(* IEC 61131-3 sources: stc/stdlib/vendor/beckhoff, 10 files *)

(* ---- common_types.st ---- *)
(* Common types used across Beckhoff TwinCAT 3 libraries *)
(* Stub declarations for stc type-checking. No implementation bodies. *)

(* AXIS_REF -- Opaque axis reference structure used by all MC_* blocks *)
TYPE AXIS_REF :
STRUCT
    NcToPlc     : DINT;
    PlcToNc     : DINT;
END_STRUCT
END_TYPE

(* MC_Direction -- Motion direction for MC_MoveAbsolute, MC_MoveVelocity *)
TYPE MC_Direction : (
    mcPositiveDirection,
    mcNegativeDirection,
    mcCurrentDirection,
    mcShortestWay
);
END_TYPE

(* T_AmsNetId -- AMS Net ID string for ADS communication *)
TYPE T_AmsNetId : STRING(23); END_TYPE

(* T_AmsPort -- AMS port number *)
TYPE T_AmsPort : UINT; END_TYPE

(* T_MaxString -- General-purpose maximum-length string *)
TYPE T_MaxString : STRING(255); END_TYPE

(* E_OpenPath -- File open path options for FB_FileOpen *)
TYPE E_OpenPath : (
    PATH_GENERIC,
    PATH_BOOTPATH,
    PATH_BOOTPRJPATH
);
END_TYPE

(* PVOID -- untyped address. TwinCAT defines PVOID as UXINT (ULINT on 64-bit,
   UDINT on 32-bit). stc declares it as POINTER TO BYTE (locked Phase 21
   decision). Phase 22 must make ADR(...) results and any POINTER TO <T>
   assignable to PVOID. *)
TYPE PVOID : POINTER TO BYTE; END_TYPE

(* Platform-width integer aliases (TwinCAT PLC manual 16.5.11), 64-bit sizes *)
TYPE __XWORD : LWORD; END_TYPE

TYPE XWORD : LWORD; END_TYPE

TYPE UXINT : ULINT; END_TYPE

TYPE __UXINT : ULINT; END_TYPE

TYPE XINT : LINT; END_TYPE

TYPE __XINT : LINT; END_TYPE

(* AMSPORT -- AMS port number (Tc2_System alias) *)
TYPE AMSPORT : UINT; END_TYPE

(* ---- tc3_ipcdiag.st ---- *)
(* Tc3_IPCDiag -- placeholder stub *)
(* No symbols from this library are used by sildarvinnsla; the file is
   present so the library reference resolves. The marker type below keeps
   the one-declaration-per-stub rule and is not a Beckhoff symbol. *)

TYPE T_Tc3IPCDiagStubMarker : BOOL; END_TYPE

(* ---- tc3_module.st ---- *)
(* Tc3_Module -- placeholder stub *)
(* No symbols from this library are used by sildarvinnsla; the file is
   present so the library reference resolves. The marker type below keeps
   the one-declaration-per-stub rule and is not a Beckhoff symbol. *)

TYPE T_Tc3ModuleStubMarker : BOOL; END_TYPE

(* ---- tc2_ethercat.st ---- *)
(* Tc2_EtherCAT -- EtherCAT diagnostics and mailbox function blocks *)
(* Stub declarations for stc type-checking. No implementation bodies. *)
(* Source: TwinCAT 3 PLC Lib Tc2_EtherCAT manual v1.10.0. *)
(* E_EcSlaveState, EcDiagParam and FB_EcDeviceDiag are deliberately NOT
   declared here: they are SVNCoreComponents declarations, not Beckhoff
   ones, and must resolve from that library. *)

TYPE E_EcAdressingType : (
    eAdressingType_AutoInc := 1,
    eAdressingType_Fixed,
    eAdressingType_Broadcast
);
END_TYPE

TYPE ST_EcSlaveState :
STRUCT
    deviceState     : BYTE;
    linkState       : BYTE;
END_STRUCT
END_TYPE

TYPE ST_EcCrcError :
STRUCT
    portA           : UDINT;
    portB           : UDINT;
    portC           : UDINT;
END_STRUCT
END_TYPE

TYPE ST_EcCrcErrorEx :
STRUCT
    portA           : UDINT;
    portB           : UDINT;
    portC           : UDINT;
    portD           : UDINT;
END_STRUCT
END_TYPE

(* Global constants, section 14.1 (subset) *)
VAR_GLOBAL CONSTANT
    EC_AMSPORT_MASTER               : UINT := 16#FFFF;
    EC_MAX_SLAVES                   : UINT := 16#FFFF;
    EC_DEVICE_STATE_MASK            : BYTE := 16#0F;
    EC_DEVICE_STATE_INIT            : BYTE := 16#01;
    EC_DEVICE_STATE_PREOP           : BYTE := 16#02;
    EC_DEVICE_STATE_BOOTSTRAP       : BYTE := 16#03;
    EC_DEVICE_STATE_SAFEOP          : BYTE := 16#04;
    EC_DEVICE_STATE_OP              : BYTE := 16#08;
    EC_DEVICE_STATE_ERROR           : BYTE := 16#10;
    EC_DEVICE_STATE_INVALID_VPRS    : BYTE := 16#20;
    EC_DEVICE_STATE_INITCMD_ERROR   : BYTE := 16#40;
    EC_LINK_STATE_OK                : BYTE := 16#00;
    EC_LINK_STATE_NOT_PRESENT       : BYTE := 16#01;
    EC_LINK_STATE_LINK_WITHOUT_COMM : BYTE := 16#02;
    EC_LINK_STATE_MISSING_LINK      : BYTE := 16#04;
    EC_LINK_STATE_ADDITIONAL_LINK   : BYTE := 16#08;
    EC_LINK_STATE_PORT_A            : BYTE := 16#10;
    EC_LINK_STATE_PORT_B            : BYTE := 16#20;
    EC_LINK_STATE_PORT_C            : BYTE := 16#40;
    EC_LINK_STATE_PORT_D            : BYTE := 16#80;
END_VAR

(* Section 3.2 *)
FUNCTION_BLOCK FB_EcPhysicalWriteCmd
VAR_INPUT
    sNetId          : T_AmsNetId;
    adp             : UINT;
    ado             : UINT;
    len             : UDINT;
    eType           : E_EcAdressingType := eAdressingType_Fixed;
    pSrcBuf         : PVOID;
    bExecute        : BOOL;
    tTimeout        : TIME := DEFAULT_ADS_TIMEOUT;
END_VAR
VAR_OUTPUT
    bBusy           : BOOL;
    bError          : BOOL;
    nErrId          : UDINT;
    wkc             : UINT;
END_VAR
END_FUNCTION_BLOCK

(* Section 4.3 *)
FUNCTION_BLOCK FB_EcGetAllSlaveAddr
VAR_INPUT
    sNetId          : T_AmsNetId;
    pAddrBuf        : POINTER TO ARRAY[0..EC_MAX_SLAVES] OF UINT;
    cbBufLen        : UDINT;
    bExecute        : BOOL;
    tTimeout        : TIME := DEFAULT_ADS_TIMEOUT;
END_VAR
VAR_OUTPUT
    bBusy           : BOOL;
    bError          : BOOL;
    nErrId          : UDINT;
    nSlaves         : UINT;
END_VAR
END_FUNCTION_BLOCK

(* Section 4.4 *)
FUNCTION_BLOCK FB_EcGetAllSlaveCrcErrors
VAR_INPUT
    sNetId          : T_AmsNetId;
    pCrcErrorBuf    : POINTER TO ARRAY[0..EC_MAX_SLAVES] OF DWORD;
    cbBufLen        : UDINT;
    bExecute        : BOOL;
    tTimeout        : TIME := DEFAULT_ADS_TIMEOUT;
END_VAR
VAR_OUTPUT
    bBusy           : BOOL;
    bError          : BOOL;
    nErrId          : UDINT;
    nSlaves         : UINT;
END_VAR
END_FUNCTION_BLOCK

(* Section 4.12 *)
FUNCTION_BLOCK FB_EcGetSlaveCrcError
VAR_INPUT
    sNetId          : T_AmsNetId;
    nSlaveAddr      : UINT;
    bExecute        : BOOL;
    tTimeout        : TIME := DEFAULT_ADS_TIMEOUT;
END_VAR
VAR_OUTPUT
    bBusy           : BOOL;
    bError          : BOOL;
    nErrId          : UDINT;
    crcError        : ST_EcCrcError;
END_VAR
END_FUNCTION_BLOCK

(* Section 4.13 (tTimeout has no default in the manual) *)
FUNCTION_BLOCK FB_EcGetSlaveCrcErrorEx
VAR_INPUT
    sNetId          : T_AmsNetId;
    nSlaveAddr      : UINT;
    bExecute        : BOOL;
    tTimeout        : TIME;
END_VAR
VAR_OUTPUT
    bBusy           : BOOL;
    bError          : BOOL;
    nErrId          : UDINT;
    CrcError        : ST_EcCrcErrorEx;
END_VAR
END_FUNCTION_BLOCK

(* Section 5.1 *)
FUNCTION_BLOCK FB_EcGetAllSlaveStates
VAR_INPUT
    sNetId          : T_AmsNetId;
    pStateBuf       : POINTER TO ARRAY[0..EC_MAX_SLAVES] OF ST_EcSlaveState;
    cbBufLen        : UDINT;
    bExecute        : BOOL;
    tTimeout        : TIME := DEFAULT_ADS_TIMEOUT;
END_VAR
VAR_OUTPUT
    bBusy           : BOOL;
    bError          : BOOL;
    nErrId          : UDINT;
    nSlaves         : UINT;
END_VAR
END_FUNCTION_BLOCK

(* Section 5.3 *)
FUNCTION_BLOCK FB_EcGetMasterState
VAR_INPUT
    sNetId          : T_AmsNetId;
    bExecute        : BOOL;
    tTimeout        : TIME := DEFAULT_ADS_TIMEOUT;
END_VAR
VAR_OUTPUT
    bBusy           : BOOL;
    bError          : BOOL;
    nErrId          : UDINT;
    state           : WORD;
END_VAR
END_FUNCTION_BLOCK

(* Section 5.4 *)
FUNCTION_BLOCK FB_EcGetSlaveState
VAR_INPUT
    sNetId          : T_AmsNetId;
    nSlaveAddr      : UINT;
    bExecute        : BOOL;
    tTimeout        : TIME := DEFAULT_ADS_TIMEOUT;
END_VAR
VAR_OUTPUT
    bBusy           : BOOL;
    bError          : BOOL;
    nErrId          : UDINT;
    state           : ST_EcSlaveState;
END_VAR
END_FUNCTION_BLOCK

(* Section 5.9 *)
FUNCTION_BLOCK FB_EcSetSlaveState
VAR_INPUT
    sNetId          : T_AmsNetId;
    nSlaveAddr      : UINT;
    bExecute        : BOOL;
    tTimeout        : TIME := T#10S;
    reqState        : WORD;
END_VAR
VAR_OUTPUT
    bBusy           : BOOL;
    bError          : BOOL;
    nErrId          : UDINT;
    currState       : ST_EcSlaveState;
END_VAR
END_FUNCTION_BLOCK

(* Section 7.1 (Beckhoff also spells it FB_EcCoeSdoRead; names are case-insensitive) *)
FUNCTION_BLOCK FB_EcCoESdoRead
VAR_INPUT
    sNetId          : T_AmsNetId;
    nSlaveAddr      : UINT;
    nSubIndex       : BYTE;
    nIndex          : WORD;
    pDstBuf         : PVOID;
    cbBufLen        : UDINT;
    bExecute        : BOOL;
    tTimeout        : TIME := DEFAULT_ADS_TIMEOUT;
END_VAR
VAR_OUTPUT
    bBusy           : BOOL;
    bError          : BOOL;
    nErrId          : UDINT;
    cbRead          : UDINT;
END_VAR
END_FUNCTION_BLOCK

(* Section 7.3 *)
FUNCTION_BLOCK FB_EcCoESdoWrite
VAR_INPUT
    sNetId          : T_AmsNetId;
    nSlaveAddr      : UINT;
    nSubIndex       : BYTE;
    nIndex          : WORD;
    pSrcBuf         : PVOID;
    cbBufLen        : UDINT;
    bExecute        : BOOL;
    tTimeout        : TIME := DEFAULT_ADS_TIMEOUT;
END_VAR
VAR_OUTPUT
    bBusy           : BOOL;
    bError          : BOOL;
    nErrId          : UDINT;
END_VAR
END_FUNCTION_BLOCK

(* ---- tc2_mc2.st ---- *)
(* Tc2_MC2 -- PLCopen Motion Control function blocks for Beckhoff TwinCAT 3 *)
(* Stub declarations for stc type-checking. No implementation bodies. *)

FUNCTION_BLOCK MC_Power
VAR_INPUT
    Axis            : AXIS_REF;
    Enable          : BOOL;
    Enable_Positive : BOOL;
    Enable_Negative : BOOL;
    Override_V      : LREAL := 100.0;
END_VAR
VAR_OUTPUT
    Status      : BOOL;
    Busy        : BOOL;
    Active      : BOOL;
    Error       : BOOL;
    ErrorID     : UDINT;
END_VAR
END_FUNCTION_BLOCK

FUNCTION_BLOCK MC_MoveAbsolute
VAR_INPUT
    Axis            : AXIS_REF;
    Execute         : BOOL;
    Position        : LREAL;
    Velocity        : LREAL;
    Acceleration    : LREAL;
    Deceleration    : LREAL;
    Jerk            : LREAL;
    Direction       : MC_Direction;
END_VAR
VAR_OUTPUT
    Done            : BOOL;
    Busy            : BOOL;
    Active          : BOOL;
    CommandAborted  : BOOL;
    Error           : BOOL;
    ErrorID         : UDINT;
END_VAR
END_FUNCTION_BLOCK

FUNCTION_BLOCK MC_MoveRelative
VAR_INPUT
    Axis            : AXIS_REF;
    Execute         : BOOL;
    Distance        : LREAL;
    Velocity        : LREAL;
    Acceleration    : LREAL;
    Deceleration    : LREAL;
    Jerk            : LREAL;
END_VAR
VAR_OUTPUT
    Done            : BOOL;
    Busy            : BOOL;
    Active          : BOOL;
    CommandAborted  : BOOL;
    Error           : BOOL;
    ErrorID         : UDINT;
END_VAR
END_FUNCTION_BLOCK

FUNCTION_BLOCK MC_MoveVelocity
VAR_INPUT
    Axis            : AXIS_REF;
    Execute         : BOOL;
    Velocity        : LREAL;
    Acceleration    : LREAL;
    Deceleration    : LREAL;
    Jerk            : LREAL;
    Direction       : MC_Direction;
END_VAR
VAR_OUTPUT
    InVelocity      : BOOL;
    Busy            : BOOL;
    Active          : BOOL;
    CommandAborted  : BOOL;
    Error           : BOOL;
    ErrorID         : UDINT;
END_VAR
END_FUNCTION_BLOCK

FUNCTION_BLOCK MC_Stop
VAR_INPUT
    Axis            : AXIS_REF;
    Execute         : BOOL;
    Deceleration    : LREAL;
    Jerk            : LREAL;
END_VAR
VAR_OUTPUT
    Done            : BOOL;
    Busy            : BOOL;
    Active          : BOOL;
    CommandAborted  : BOOL;
    Error           : BOOL;
    ErrorID         : UDINT;
END_VAR
END_FUNCTION_BLOCK

FUNCTION_BLOCK MC_Home
VAR_INPUT
    Axis            : AXIS_REF;
    Execute         : BOOL;
    Position        : LREAL;
END_VAR
VAR_OUTPUT
    Done            : BOOL;
    Busy            : BOOL;
    Active          : BOOL;
    CommandAborted  : BOOL;
    Error           : BOOL;
    ErrorID         : UDINT;
END_VAR
END_FUNCTION_BLOCK

FUNCTION_BLOCK MC_Reset
VAR_INPUT
    Axis            : AXIS_REF;
    Execute         : BOOL;
END_VAR
VAR_OUTPUT
    Done            : BOOL;
    Busy            : BOOL;
    Error           : BOOL;
    ErrorID         : UDINT;
END_VAR
END_FUNCTION_BLOCK

FUNCTION_BLOCK MC_ReadActualPosition
VAR_INPUT
    Axis            : AXIS_REF;
    Enable          : BOOL;
END_VAR
VAR_OUTPUT
    Valid           : BOOL;
    Busy            : BOOL;
    Error           : BOOL;
    ErrorID         : UDINT;
    Position        : LREAL;
END_VAR
END_FUNCTION_BLOCK

FUNCTION_BLOCK MC_ReadActualVelocity
VAR_INPUT
    Axis            : AXIS_REF;
    Enable          : BOOL;
END_VAR
VAR_OUTPUT
    Valid           : BOOL;
    Busy            : BOOL;
    Error           : BOOL;
    ErrorID         : UDINT;
    ActualVelocity  : LREAL;
END_VAR
END_FUNCTION_BLOCK

FUNCTION_BLOCK MC_ReadStatus
VAR_INPUT
    Axis            : AXIS_REF;
    Enable          : BOOL;
END_VAR
VAR_OUTPUT
    Valid               : BOOL;
    Busy                : BOOL;
    Error               : BOOL;
    ErrorID             : UDINT;
    ErrorStop           : BOOL;
    Disabled            : BOOL;
    Stopping            : BOOL;
    StandStill          : BOOL;
    DiscreteMotion      : BOOL;
    ContinuousMotion    : BOOL;
    SynchronizedMotion  : BOOL;
    Homing              : BOOL;
END_VAR
END_FUNCTION_BLOCK

(* ---- tc2_modbussrv.st ---- *)
(* Tc2_ModbusSrv -- Modbus TCP client function blocks (TF6250) *)
(* Stub declarations for stc type-checking. No implementation bodies. *)
(* Source: TF6250 TC3 Modbus TCP manual section 6.1.2. Section 6.1 states the
   Modbus functions are implemented in the PLC library Tc2_ModbusSrv, which is
   the library name TwinCAT projects reference, so the client FBs live here. *)

VAR_GLOBAL CONSTANT
    MODBUS_TCP_PORT : UINT := 502;      (* value assumed: Modbus TCP standard port *)
END_VAR

(* Modbus function 1 *)
FUNCTION_BLOCK FB_MBReadCoils
VAR_INPUT
    sIPAddr         : STRING(15);
    nTCPPort        : UINT := MODBUS_TCP_PORT;
    nUnitID         : BYTE := 16#FF;
    nQuantity       : WORD;
    nMBAddr         : WORD;
    cbLength        : UDINT;
    pDestAddr       : POINTER TO BYTE;
    bExecute        : BOOL;
    tTimeout        : TIME;
END_VAR
VAR_OUTPUT
    bBUSY           : BOOL;
    bError          : BOOL;
    nErrId          : UDINT;
    cbRead          : UDINT;
END_VAR
END_FUNCTION_BLOCK

(* Modbus function 2 *)
FUNCTION_BLOCK FB_MBReadInputs
VAR_INPUT
    sIPAddr         : STRING(15);
    nTCPPort        : UINT := MODBUS_TCP_PORT;
    nUnitID         : BYTE := 16#FF;
    nQuantity       : WORD;
    nMBAddr         : WORD;
    cbLength        : UDINT;
    pDestAddr       : POINTER TO BYTE;
    bExecute        : BOOL;
    tTimeout        : TIME;
END_VAR
VAR_OUTPUT
    bBUSY           : BOOL;
    bError          : BOOL;
    nErrId          : UDINT;
    cbRead          : UDINT;
END_VAR
END_FUNCTION_BLOCK

(* Modbus function 3 *)
FUNCTION_BLOCK FB_MBReadRegs
VAR_INPUT
    sIPAddr         : STRING(15);
    nTCPPort        : UINT := MODBUS_TCP_PORT;
    nUnitID         : BYTE := 16#FF;
    nQuantity       : WORD;
    nMBAddr         : WORD;
    cbLength        : UDINT;
    pDestAddr       : POINTER TO BYTE;
    bExecute        : BOOL;
    tTimeout        : TIME;
END_VAR
VAR_OUTPUT
    bBUSY           : BOOL;
    bError          : BOOL;
    nErrId          : UDINT;
    cbRead          : UDINT;
END_VAR
END_FUNCTION_BLOCK

(* Modbus function 4 *)
FUNCTION_BLOCK FB_MBReadInputRegs
VAR_INPUT
    sIPAddr         : STRING(15);
    nTCPPort        : UINT := MODBUS_TCP_PORT;
    nUnitID         : BYTE := 16#FF;
    nQuantity       : WORD;
    nMBAddr         : WORD;
    cbLength        : UDINT;
    pDestAddr       : POINTER TO BYTE;
    bExecute        : BOOL;
    tTimeout        : TIME;
END_VAR
VAR_OUTPUT
    bBUSY           : BOOL;
    bError          : BOOL;
    nErrId          : UDINT;
    cbRead          : UDINT;
END_VAR
END_FUNCTION_BLOCK

(* Modbus function 5 *)
FUNCTION_BLOCK FB_MBWriteSingleCoil
VAR_INPUT
    sIPAddr         : STRING(15);
    nTCPPort        : UINT := MODBUS_TCP_PORT;
    nUnitID         : BYTE := 16#FF;
    nMBAddr         : WORD;
    nValue          : WORD;
    bExecute        : BOOL;
    tTimeout        : TIME;
END_VAR
VAR_OUTPUT
    bBUSY           : BOOL;
    bError          : BOOL;
    nErrId          : UDINT;
END_VAR
END_FUNCTION_BLOCK

(* Modbus function 6 *)
FUNCTION_BLOCK FB_MBWriteSingleReg
VAR_INPUT
    sIPAddr         : STRING(15);
    nTCPPort        : UINT := MODBUS_TCP_PORT;
    nUnitID         : BYTE := 16#FF;
    nMBAddr         : WORD;
    nValue          : WORD;
    bExecute        : BOOL;
    tTimeout        : TIME;
END_VAR
VAR_OUTPUT
    bBUSY           : BOOL;
    bError          : BOOL;
    nErrId          : UDINT;
END_VAR
END_FUNCTION_BLOCK

(* Modbus function 15 *)
FUNCTION_BLOCK FB_MBWriteCoils
VAR_INPUT
    sIPAddr         : STRING(15);
    nTCPPort        : UINT := MODBUS_TCP_PORT;
    nUnitID         : BYTE := 16#FF;
    nQuantity       : WORD;
    nMBAddr         : WORD;
    cbLength        : UDINT;
    pSrcAddr        : POINTER TO BYTE;
    bExecute        : BOOL;
    tTimeout        : TIME;
END_VAR
VAR_OUTPUT
    bBUSY           : BOOL;
    bError          : BOOL;
    nErrId          : UDINT;
END_VAR
END_FUNCTION_BLOCK

(* Modbus function 16 *)
FUNCTION_BLOCK FB_MBWriteRegs
VAR_INPUT
    sIPAddr         : STRING(15);
    nTCPPort        : UINT := MODBUS_TCP_PORT;
    nUnitID         : BYTE := 16#FF;
    nQuantity       : WORD;
    nMBAddr         : WORD;
    cbLength        : UDINT;
    pSrcAddr        : POINTER TO BYTE;
    bExecute        : BOOL;
    tTimeout        : TIME;
END_VAR
VAR_OUTPUT
    bBUSY           : BOOL;
    bError          : BOOL;
    nErrId          : UDINT;
END_VAR
END_FUNCTION_BLOCK

(* Modbus function 23 *)
FUNCTION_BLOCK FB_MBReadWriteRegs
VAR_INPUT
    sIPAddr         : STRING(15);
    nTCPPort        : UINT := MODBUS_TCP_PORT;
    nUnitID         : BYTE := 16#FF;
    nReadQuantity   : WORD;
    nMBReadAddr     : WORD;
    nWriteQuantity  : WORD;
    nMBWriteAddr    : WORD;
    cbDestLength    : UDINT;
    pDestAddr       : POINTER TO BYTE;
    cbSrcLength     : UDINT;
    pSrcAddr        : POINTER TO BYTE;
    bExecute        : BOOL;
    tTimeout        : TIME;
END_VAR
VAR_OUTPUT
    bBUSY           : BOOL;
    bError          : BOOL;
    nErrId          : UDINT;
    cbRead          : UDINT;
END_VAR
END_FUNCTION_BLOCK

(* ---- tc2_serialcom.st ---- *)
(* Tc2_SerialCom -- serial communication function blocks (TF6340) *)
(* Stub declarations for stc type-checking. No implementation bodies. *)
(* Source: TF6340 TC3 Serial Communication manual section 5. The real type
   names are ComBuffer, ComSerialLineMode_t and ComError_t (ST_ComBuffer and
   E_ComMode do not exist). At the time of writing no plcproj-listed
   sildarvinnsla source uses these names (only Baader/PLC-TASK.md mentions
   them) and Baader does not reference Tc2_SerialCom; this stub is exercised
   by the committed usage fixture only. *)

TYPE ComBuffer :
STRUCT
    Buffer          : ARRAY[0..300] OF BYTE;
    RdIdx           : INT;
    WrIdx           : INT;
    Count           : INT;
    FreeByte        : INT;
    Error           : INT;
    blocked         : BOOL;
END_STRUCT
END_TYPE

TYPE ComSerialLineMode_t : (
    SERIALLINEMODE_DEFAULT,
    SERIALLINEMODE_KL6_3B_ALTERNATIVE,
    SERIALLINEMODE_KL6_5B_STANDARD,
    SERIALLINEMODE_KL6_22B_STANDARD,
    SERIALLINEMODE_PC_COM_PORT,
    SERIALLINEMODE_EL6_22B,
    SERIALLINEMODE_IE6_11B
);
END_TYPE

TYPE ComError_t : (
    COMERROR_NOERROR := 0,
    COMERROR_PARAMETERCHANGED := 1,
    COMERROR_TXBUFFOVERRUN := 2,
    COMERROR_STRINGOVERRUN := 10,
    COMERROR_ZEROCHARINVALID := 11,
    COMERROR_INVALIDPOINTER := 20,
    COMERROR_INVALIDRXPOINTER := 21,
    COMERROR_INVALIDRXLENGTH := 22,
    COMERROR_DATASIZEOVERRUN := 23,
    COMERROR_INVALIDPROCESSDATASIZE := 24,
    COMERROR_MODENOTSUPPORTED := 16#0101,
    COMERROR_INVALIDCHANNELNUMBER := 16#0102,
    COMERROR_INVALIDBAUDRATE := 16#1001,
    COMERROR_INVALIDNUMDATABITS := 16#1002,
    COMERROR_INVALIDNUMSTOPBITS := 16#1003,
    COMERROR_INVALIDPARITY := 16#1004,
    COMERROR_INVALIDHANDSHAKE := 16#1005,
    COMERROR_INVALIDNUMREGISTERS := 16#1006,
    COMERROR_INVALIDREGISTER := 16#1007,
    COMERROR_TIMEOUT := 16#1008
);
END_TYPE

(* Section 5 *)
FUNCTION_BLOCK SerialLineControl
VAR_INPUT
    Mode            : ComSerialLineMode_t;
    pComIn          : POINTER TO BYTE;
    pComOut         : POINTER TO BYTE;
    SizeComIn       : INT;
END_VAR
VAR_IN_OUT
    TxBuffer        : ComBuffer;
    RxBuffer        : ComBuffer;
END_VAR
VAR_OUTPUT
    Error           : BOOL;
    ErrorID         : ComError_t;
END_VAR
END_FUNCTION_BLOCK

(* Section 5 *)
FUNCTION_BLOCK SendByte
VAR_INPUT
    SendByte        : BYTE;
END_VAR
VAR_IN_OUT
    TxBuffer        : ComBuffer;
END_VAR
VAR_OUTPUT
    Busy            : BOOL;
    Error           : ComError_t;
END_VAR
END_FUNCTION_BLOCK

(* Section 5 *)
FUNCTION_BLOCK SendString
VAR_INPUT
    SendString      : STRING;
END_VAR
VAR_IN_OUT
    TxBuffer        : ComBuffer;
END_VAR
VAR_OUTPUT
    Busy            : BOOL;
    Error           : ComError_t;
END_VAR
END_FUNCTION_BLOCK

(* Section 5 *)
FUNCTION_BLOCK ReceiveByte
VAR_IN_OUT
    RXBuffer        : ComBuffer;
END_VAR
VAR_OUTPUT
    ByteReceived    : BOOL;
    ReceivedByte    : BYTE;
    Error           : ComError_t;
END_VAR
END_FUNCTION_BLOCK

(* Section 5 *)
FUNCTION_BLOCK ReceiveString
VAR_INPUT
    Prefix          : STRING;
    Suffix          : STRING;
    Timeout         : TIME;
    Reset           : BOOL;
END_VAR
VAR_IN_OUT
    ReceivedString  : STRING;
    RXBuffer        : ComBuffer;
END_VAR
VAR_OUTPUT
    StringReceived  : BOOL;
    busy            : BOOL;
    Error           : ComError_t;
    RxTimeout       : BOOL;
END_VAR
END_FUNCTION_BLOCK

(* Section 5 *)
FUNCTION_BLOCK ClearComBuffer
VAR_IN_OUT
    Buffer          : ComBuffer;
END_VAR
END_FUNCTION_BLOCK

(* ---- tc2_system.st ---- *)
(* Tc2_System -- System function blocks for Beckhoff TwinCAT 3 *)
(* Stub declarations for stc type-checking. No implementation bodies. *)
(* RTC is declared by Beckhoff in Tc2_Utilities (manual v2.18.2 section 3.79).
   It lives here because Tc2_Standard is built in to stc, and every stub
   closure includes tc2_system, so a project referencing only Tc2_Standard
   and Tc2_System still resolves RTC. *)

(* T_AmsNetIdArr -- AMS Net ID as six bytes (section 5, BYTE not USINT) *)
TYPE T_AmsNetIdArr : ARRAY[0..5] OF BYTE; END_TYPE

(* AMSNETID -- AMS Net ID byte array (TwinCAT type system, 6 x BYTE) *)
TYPE AMSNETID : ARRAY[0..5] OF BYTE; END_TYPE

(* AMSADDR -- AMS address; port is WORD in the TwinCAT type system *)
TYPE AMSADDR :
STRUCT
    netId       : AMSNETID;
    port        : WORD;
END_STRUCT
END_TYPE

(* ST_AmsAddr -- AMS address (section 5.11) *)
TYPE ST_AmsAddr :
STRUCT
    netId       : T_AmsNetIdArr;
    port        : T_AmsPort;
END_STRUCT
END_TYPE

VAR_GLOBAL CONSTANT
    DEFAULT_ADS_TIMEOUT : TIME := T#5S;     (* name cited; value assumed *)
    MAX_STRING_LENGTH   : UDINT := 255;     (* section 5.20 *)
END_VAR

(* F_CreateAmsNetId -- byte array to dotted Net ID string (section 4.2.4) *)
FUNCTION F_CreateAmsNetId : T_AmsNetId
VAR_INPUT
    nIds        : T_AmsNetIdArr;
END_VAR
END_FUNCTION

(* RTC -- software real-time clock (Tc2_Utilities section 3.79, see header) *)
FUNCTION_BLOCK RTC
VAR_INPUT
    EN          : BOOL;
    PDT         : DATE_AND_TIME;
END_VAR
VAR_OUTPUT
    Q           : BOOL;
    CDT         : DATE_AND_TIME;
END_VAR
END_FUNCTION_BLOCK

FUNCTION_BLOCK ADSREAD
VAR_INPUT
    NETID       : T_AmsNetId;
    PORT        : T_AmsPort;
    IDXGRP      : UDINT;
    IDXOFFS     : UDINT;
    LEN         : UDINT;
    DESTADDR    : PVOID;
    READ        : BOOL;
    TMOUT       : TIME := DEFAULT_ADS_TIMEOUT;
END_VAR
VAR_OUTPUT
    BUSY        : BOOL;
    ERR         : BOOL;
    ERRID       : UDINT;
END_VAR
END_FUNCTION_BLOCK

FUNCTION_BLOCK ADSWRITE
VAR_INPUT
    NETID       : T_AmsNetId;
    PORT        : T_AmsPort;
    IDXGRP      : UDINT;
    IDXOFFS     : UDINT;
    LEN         : UDINT;
    SRCADDR     : PVOID;
    WRITE       : BOOL;
    TMOUT       : TIME := DEFAULT_ADS_TIMEOUT;
END_VAR
VAR_OUTPUT
    BUSY        : BOOL;
    ERR         : BOOL;
    ERRID       : UDINT;
END_VAR
END_FUNCTION_BLOCK

FUNCTION_BLOCK FB_FileOpen
VAR_INPUT
    sNetId      : T_AmsNetId;
    sPathName   : T_MaxString;
    nMode       : DWORD;
    ePath       : E_OpenPath := PATH_GENERIC;
    bExecute    : BOOL;
    tTimeout    : TIME := T#5S;
END_VAR
VAR_OUTPUT
    bBusy       : BOOL;
    bError      : BOOL;
    nErrId      : UDINT;
    hFile       : UINT;
END_VAR
END_FUNCTION_BLOCK

FUNCTION_BLOCK FB_FileClose
VAR_INPUT
    sNetId      : T_AmsNetId;
    hFile       : UINT;
    bExecute    : BOOL;
    tTimeout    : TIME := T#5S;
END_VAR
VAR_OUTPUT
    bBusy       : BOOL;
    bError      : BOOL;
    nErrId      : UDINT;
END_VAR
END_FUNCTION_BLOCK

FUNCTION_BLOCK FB_FileRead
VAR_INPUT
    sNetId      : T_AmsNetId;
    hFile       : UINT;
    pReadBuff   : UDINT;
    cbReadLen   : UDINT;
    bExecute    : BOOL;
    tTimeout    : TIME := T#5S;
END_VAR
VAR_OUTPUT
    bBusy       : BOOL;
    bError      : BOOL;
    nErrId      : UDINT;
    cbRead      : UDINT;
    bEOF        : BOOL;
END_VAR
END_FUNCTION_BLOCK

FUNCTION_BLOCK FB_FileWrite
VAR_INPUT
    sNetId      : T_AmsNetId;
    hFile       : UINT;
    pWriteBuff  : UDINT;
    cbWriteLen  : UDINT;
    bExecute    : BOOL;
    tTimeout    : TIME := T#5S;
END_VAR
VAR_OUTPUT
    bBusy       : BOOL;
    bError      : BOOL;
    nErrId      : UDINT;
    cbWrite     : UDINT;
END_VAR
END_FUNCTION_BLOCK

FUNCTION MEMCPY : UDINT
VAR_INPUT
    destAddr    : PVOID;
    srcAddr     : PVOID;
    n           : UDINT;
END_VAR
END_FUNCTION

FUNCTION MEMSET : UDINT
VAR_INPUT
    destAddr    : PVOID;
    fillByte    : USINT;
    n           : UDINT;
END_VAR
END_FUNCTION

FUNCTION MEMMOVE : UDINT
VAR_INPUT
    destAddr    : PVOID;
    srcAddr     : PVOID;
    n           : UDINT;
END_VAR
END_FUNCTION

FUNCTION MEMCMP : DINT
VAR_INPUT
    pBuf1       : PVOID;
    pBuf2       : PVOID;
    n           : UDINT;
END_VAR
END_FUNCTION

(* ---- tc2_utilities.st ---- *)
(* Tc2_Utilities -- Utility function blocks for Beckhoff TwinCAT 3 *)
(* Stub declarations for stc type-checking. No implementation bodies. *)

FUNCTION_BLOCK FB_FormatString
VAR_INPUT
    sFormat     : T_MaxString;
    arg1        : T_MaxString;
    arg2        : T_MaxString;
    arg3        : T_MaxString;
    arg4        : T_MaxString;
    arg5        : T_MaxString;
    arg6        : T_MaxString;
    arg7        : T_MaxString;
    arg8        : T_MaxString;
    arg9        : T_MaxString;
    arg10       : T_MaxString;
    bExecute    : BOOL;
END_VAR
VAR_OUTPUT
    bDone       : BOOL;
    bError      : BOOL;
    nErrId      : UDINT;
    sOut        : T_MaxString;
END_VAR
END_FUNCTION_BLOCK

FUNCTION CRC16 : UINT
VAR_INPUT
    pData       : UDINT;
    cbLen       : UDINT;
    nInit       : UINT;
    nPoly       : UINT;
END_VAR
END_FUNCTION

FUNCTION CRC32 : UDINT
VAR_INPUT
    pData       : UDINT;
    cbLen       : UDINT;
    nInit       : UDINT;
    nPoly       : UDINT;
END_VAR
END_FUNCTION

(* TIMESTRUCT -- Windows SYSTEMTIME layout *)
TYPE TIMESTRUCT :
STRUCT
    wYear           : WORD;
    wMonth          : WORD;
    wDayOfWeek      : WORD;
    wDay            : WORD;
    wHour           : WORD;
    wMinute         : WORD;
    wSecond         : WORD;
    wMilliseconds   : WORD;
END_STRUCT
END_TYPE

(* E_TimeZoneID -- time zone state reported by FB_LocalSystemTime *)
TYPE E_TimeZoneID : (
    eTimeZoneID_Invalid := -1,
    eTimeZoneID_Unknown := 0,
    eTimeZoneID_Standard := 1,
    eTimeZoneID_Daylight := 2
);
END_TYPE

(* FB_LocalSystemTime -- local Windows time, synchronised cyclically (3.47) *)
FUNCTION_BLOCK FB_LocalSystemTime
VAR_INPUT
    sNetID      : T_AmsNetId := '';
    bEnable     : BOOL;
    dwCycle     : DWORD(1..86400) := 5;
    dwOpt       : DWORD := 1;
    tTimeout    : TIME := DEFAULT_ADS_TIMEOUT;
END_VAR
VAR_OUTPUT
    bValid      : BOOL;
    systemTime  : TIMESTRUCT;
    tzID        : E_TimeZoneID := eTimeZoneID_Invalid;
END_VAR
END_FUNCTION_BLOCK

(* SYSTEMTIME_TO_DT -- TIMESTRUCT to DATE_AND_TIME (4.1.18) *)
FUNCTION SYSTEMTIME_TO_DT : DT
VAR_INPUT
    TIMESTR     : TIMESTRUCT;
END_VAR
END_FUNCTION

(* ---- tc3_eventlogger.st ---- *)
(* Tc3_EventLogger -- Event logging for Beckhoff TwinCAT 3 *)
(* Stub declarations for stc type-checking. No implementation bodies. *)

FUNCTION_BLOCK FB_TcEventLogger
VAR_INPUT
    bExecute    : BOOL;
    nEventId    : UDINT;
    eSeverity   : INT;
    sMessage    : T_MaxString;
END_VAR
VAR_OUTPUT
    bDone       : BOOL;
    bBusy       : BOOL;
    bError      : BOOL;
    nErrId      : UDINT;
END_VAR
END_FUNCTION_BLOCK

FUNCTION_BLOCK FB_TcAlarm
VAR_INPUT
    bExecute    : BOOL;
    nEventId    : UDINT;
    eSeverity   : INT;
    sMessage    : T_MaxString;
    bConfirm    : BOOL;
    bReset      : BOOL;
END_VAR
VAR_OUTPUT
    bDone       : BOOL;
    bBusy       : BOOL;
    bError      : BOOL;
    nErrId      : UDINT;
    bActive     : BOOL;
    bConfirmed  : BOOL;
END_VAR
END_FUNCTION_BLOCK
